Yaskawa INFORM job: SUBPICK.JBI

/JOB
//NAME SUBPICK
//POS
///NPOS 1,0,0,0,0,0
///TOOL 1
///POSTYPE BASE
///RECTAN
///RCONF 0,0,0,0,0,0,0,0
C00000=674.300,134.999,685.980,-66.22,8.38,-107.67
//INST
///DATE 2026/10/26 01:18
///COMM Generated using RoboDK
///ATTR SC,RW,RJ
///GROUP1 RB1
NOP
MOVL C00000 V=300.0 ACC=100 DEC=100
DOUT OT#(7) ON
END
